// TIA Portal V20 export
Screen "Pop-up_PN_DEV_DIAG_LEGEND_Popup"  430x552
  ScreenItem "Background" at 0,0 size 430x552  Type=HmiRectangle
  ScreenItem "Text_Legend1" at 1,1 size 428x25  Type=HmiTextBox
  ScreenItem "Text_Symbol_PN-DEV_NoName" at 10,204 size 170x20  Type=HmiTextBox
  ScreenItem "Text_Symbol_PN-DEV_OK" at 10,29 size 170x20  Type=HmiTextBox
  ScreenItem "Text_Symbol_PN-DEV_Faulty" at 10,109 size 170x20  Type=HmiTextBox
  ScreenItem "Text_Symbol_PN-DEV_NotPresent" at 10,64 size 170x20  Type=HmiTextBox
  ScreenItem "Text_Symbol_PN-DEV_Deaktivated" at 10,86 size 170x20  Type=HmiTextBox
  ScreenItem "Text_PN-DEV_NoName" at 185,199 size 235x35  Type=HmiTextBox
  ScreenItem "Text_PN-DEV_OK" at 185,26 size 155x39  Type=HmiTextBox
  ScreenItem "Text_PN-DEV_Faulty" at 185,111 size 235x20  Type=HmiTextBox
  ScreenItem "Text_PN-DEV_Deaktivated" at 185,89 size 235x20  Type=HmiTextBox
  ScreenItem "Text_Legend2" at 10,365 size 120x20  Type=HmiTextBox
  ScreenItem "Cancel Mode" at 339,1 size 90x60  Type=HmiButton
  ScreenItem "Text_PN-DEV_NotPresent" at 185,67 size 235x20  Type=HmiTextBox
  ScreenItem "Text_Symbol_PN-DEV_WasFaulty" at 10,131 size 170x20  Type=HmiTextBox
  ScreenItem "Text_PN-DEV_WasFaulty" at 185,133 size 235x20  Type=HmiTextBox
  ScreenItem "Text_Symbol_PN-DEV_Problem" at 10,154 size 170x20  Type=HmiTextBox
  ScreenItem "Text_PN-DEV_Problem" at 185,155 size 235x20  Type=HmiTextBox
  ScreenItem "Text_Symbol_PN-DEV_WasProblem" at 10,176 size 170x20  Type=HmiTextBox
  ScreenItem "Text_PN-DEV_WasProblem" at 185,177 size 235x20  Type=HmiTextBox
  ScreenItem "Text_Symbol_DevNo" at 10,236 size 34x20  Type=HmiTextBox
  ScreenItem "Text_DevNo" at 49,236 size 140x20  Type=HmiTextBox
  ScreenItem "Text_SubordinateMoldulError" at 49,258 size 140x20  Type=HmiTextBox
  ScreenItem "Symbol_Tec-Unit_Type" at 185,239 size 74x16  Type=HmiTextBox
  ScreenItem "Symbol_MLFB" at 8,327 size 62x20  Type=HmiTextBox
  ScreenItem "Text_MLFB" at 75,327 size 350x35  Type=HmiTextBox
  ScreenItem "Button_Reset" at 10,387 size 60x40  Type=HmiTextBox
  ScreenItem "Button_ResetText" at 75,379 size 347x56  Type=HmiTextBox
  ScreenItem "Button_ReadNew" at 10,440 size 60x40  Type=HmiTextBox
  ScreenItem "Button_ResetText_1" at 75,435 size 347x55  Type=HmiTextBox
  ScreenItem "Button_ReadNew_1" at 10,493 size 60x40  Type=HmiTextBox
  ScreenItem "Button_ResetText_2" at 75,490 size 347x55  Type=HmiTextBox
  ScreenItem "Grafikanzeige_1" at 10,261 size 14x14  Type=HmiGraphicView
  ScreenItem "PN-Line_Vertical" at 182,266 size 100x0  Type=HmiLine
  ScreenItem "Text_SubordinateMoldulError_1" at 49,280 size 140x20  Type=HmiTextBox
  ScreenItem "Text_SubordinateMoldulError_2" at 49,302 size 140x20  Type=HmiTextBox
  ScreenItem "Text_PN-DEV_NoName_1" at 303,287 size 74x18  Type=HmiTextBox
  ScreenItem "Grafikanzeige_4" at 10,283 size 14x14  Type=HmiGraphicView
  ScreenItem "Grafikanzeige_2" at 10,305 size 14x14  Type=HmiGraphicView
  ScreenItem "Text_PN-DEV_NoName_2" at 303,258 size 108x18  Type=HmiTextBox
  ScreenItem "PN-Line_Vertical_1" at 182,297 size 100x0  Type=HmiLine
